ADAPTER pusher_info (* Adapter Interface *)
  (* Standard: 61499-1 *)
  (* Version 0.0, 10/22/2026, macie, Schneider Electric *)
  PACKAGE Main;
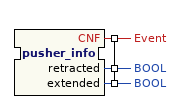
  EVENT_OUTPUT
    CNF WITH retracted, extended; (* Confirmation from Plug *)
  END_EVENT
  VAR_OUTPUT
    retracted : BOOL; (* Confirmation Data from Plug *)
    extended : BOOL; (* Indication Data from Plug *)
  END_VAR
  SERVICE SOCKET/PLUG
    SEQUENCE request_confirm
      SOCKET.REQ(REQD) -> PLUG.REQ(REQD);
      PLUG.CNF(retracted) -> SOCKET.CNF(retracted);
    END_SEQUENCE
    SEQUENCE indication_response
      PLUG.IND(extended) -> SOCKET.IND(extended);
      SOCKET.RSP(RSPD) -> PLUG.RSP(RSPD);
    END_SEQUENCE
  END_SERVICE
END_ADAPTER
